(* IEC 61131-3 sources: codesys/project-view/Device/Plc Logic/Application/000-模组/本项目/00-文件读写/字符串处理, 4 files *)

(* ---- FUN_CheckString.st ---- *)
//利用起始符和终止符，检查字符串是否完整
FUNCTION FUN_CheckString : STRING
VAR_INPUT
	RcvStr					: STRING(GlobFile.iStringLen);
	StartStr				: STRING:=GlobFile.sStartCharacter;
	EndStr					: STRING:=GlobFile.sTerminator;
END_VAR

VAR_OUTPUT
	xFromStr				: STRING(GlobFile.iStringLen);
END_VAR

VAR
	iFind_startStr			: INT;
	iFind_endStr			: INT;
	sMid					: STRING;
    suiMid					: UINT;

END_VAR
// --- implementation ---
//查找字符 StartStr
iFind_startStr:=stu.StrFindA(pst1 := ADR(RcvStr), pst2 := ADR(startStr), uiSearchStart := 1);
//查找字符 EndStr
iFind_endStr:=stu.StrFindA(pst1 := ADR(RcvStr), pst2 := ADR(endStr), uiSearchStart := 1);

IF iFind_startStr>0 AND iFind_endStr>0 THEN
	//截取字符串 '^'~'#'
	stu.StrMidA(pst := ADR(RcvStr), uiInputBufferSize := SIZEOF(ADR(RcvStr)), iLength := iFind_endStr-iFind_startStr+1, iPosition := 1 , pstResult := ADR(xFromStr), uiResultBufferSize := suiMid);

	FUN_CheckString := 'OK';

ELSE
	FUN_CheckString := 'Incomplete';//数据报文不完整

END_IF
END_FUNCTION

(* ---- FUN_CutString.st ---- *)
//根据起始符和终止符，裁剪分成字符串数组[0.199]
FUNCTION FUN_CutString : STRING
VAR_INPUT
	sString							: STRING(GlobFile.iStringLen);
	sStartCharacter					: STRING:='/';//起始符
	sTerminator						: STRING:=';';//终止符
END_VAR

VAR_OUTPUT
	asParaNum							: ARRAY[0..GlobFile.iParaLen] OF STRING;
END_VAR

VAR
	i								: UINT;
	temp							: INT;		//查找的起始位置
	iFindStartCharacter				: INT;		//查找起始符的位置
	iFindTerminator					: INT;		//查找终止符的位置

END_VAR
// --- implementation ---
(**********************************************************
例如：
sString := '/a := 123;$R$N/b := 456;';

输出：
asPara[0] => '/a := 123;'		asPara[1] => '/b := 456;'
**********************************************************)

// iFindStartCharacter := 0;
// iFindTerminator := 0;
// temp:=0;
FOR i:=0 TO GlobFile.iParaLen DO
	iFindStartCharacter := StrFindA(pst1 := ADR(sString), pst2 := ADR(sStartCharacter), uiSearchStart := INT_TO_UINT(temp+1));
	iFindTerminator := StrFindA(pst1 := ADR(sString), pst2 := ADR(sTerminator), uiSearchStart := INT_TO_UINT(temp+1));

	IF iFindStartCharacter>0 AND iFindTerminator>0 THEN	//有数据才记录下来，读到空数据就跳出循环
		StrMidA(pst := ADR(sString), uiInputBufferSize := SIZEOF(ADR(sString)), iLength := iFindTerminator-iFindStartCharacter+1, iPosition := iFindStartCharacter , pstResult := ADR(asParaNum[i]), uiResultBufferSize := 0);

		temp := iFindTerminator;//记录本次终止符的位置，下次从此位置开始搜索字符串
		iFindStartCharacter := 0;
		iFindTerminator := 0;

	ELSE
		EXIT;
	END_IF

END_FOR
END_FUNCTION

(* ---- FUN_FileStringConcat.st ---- *)
//[0..199]的数组中每个元素都连接成'/[x] := num;'
FUNCTION FUN_FileStringConcat : BOOL
VAR_INPUT
	asPara						: ARRAY[0..GlobFile.iParaLen] OF STRING;
	arNum						: ARRAY[0..GlobFile.iParaLen] OF REAL;
END_VAR

VAR_OUTPUT
	asParaNum					: ARRAY[0..GlobFile.iParaLen] OF STRING;
END_VAR

VAR
	sTmp						: STRING;
	sTmpNum						: ARRAY[0..GlobFile.iParaLen] OF STRING;
	i							: UINT;

END_VAR
// --- implementation ---
(*********************************************************
例如：
asPara[0] := 'Example';			asNum[0] := 1234;

输出：
asParaNum[0] => '/Example := 1234;' 	//有数据
asParaNum[1] => '/ := 0;' 				//没数据，即 GlobFile.sNullPara
**********************************************************)

//先把数据转成string
FOR i := 0 TO TO_UINT(GlobFile.iParaLen) DO
	sTmpNum[i] := TO_STRING(arNum[i]);
END_FOR

FOR i := 0 TO TO_UINT(GlobFile.iParaLen) DO
	IF asPara[i] = '' THEN		//如果是空字符串，就退出循环不连接
		EXIT;
	ELSE
		sTmp := CONCAT(STR1:='/' , STR2:=asPara[i] );
		sTmp := CONCAT(STR1:=sTmp , STR2:=' := ' );
		sTmp := CONCAT(STR1:=sTmp , STR2:=sTmpNum[i] );
		asParaNum[i] := CONCAT(STR1:=sTmp , STR2:=';' );
	END_IF

END_FOR
END_FUNCTION

(* ---- FUN_FindString.st ---- *)
//取str1与str2的中间字符串
FUNCTION FUN_FindString : STRING
VAR_INPUT
	str:STRING(255);		//
	str1:STRING;	//first find string
	str2:STRING;	//second find string
END_VAR

VAR
	temp1:INT;
	temp2:INT;
END_VAR
// --- implementation ---
temp1:=find(str,str1);
temp2:=find(str,str2);
FUN_FindString:=mid(str,temp2-temp1-len(str1),temp1+len(str1));	//取str1与str2的中间字符串
END_FUNCTION
